ABB RAPID module: TurnProg.mod

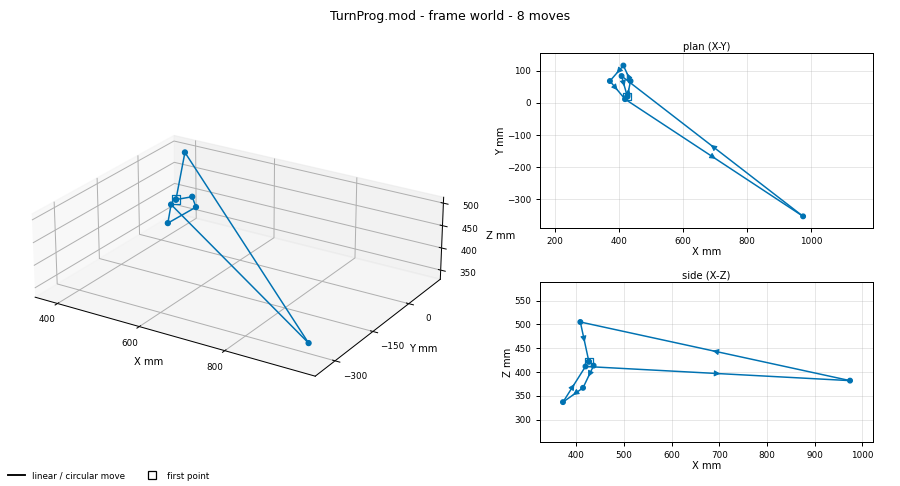
[picture p0: tool path of TurnProg.mod in frame world, 8 of 9 moves have a stored position in this frame; points joined in program order, loops and branches not executed]
%%%
  VERSION:1
  LANGUAGE:ENGLISH
%%%
MODULE MOD_TurnProg

    ! -------------------------------
    ! Define customized variables here
    ! ...

	! Tool variables:
	PERS tooldata ToolS := [TRUE,[[10.000,20.000,150.000],[1.00000000,0.00000000,0.00000000,0.00000000]],[1,[0,0,20],[1,0,0,0],0,0,0.005]];

	! Reference variables:
	PERS wobjdata FrameS := [FALSE, TRUE, "", [[0,0,0],[1,0,0,0]],[[1234.570,-98.765,50.500],[0.96592583,0.00000000,0.00000000,0.25881905]]];

	PROC Main()
		ConfJ \On;
		ConfL \Off;
		! Program generated by RoboDK v6.0.7 for ABB IRB 260 on XX/XX/XXXX 18:00:00
		! Using nominal kinematics.
		MoveL [[-640.584,506.980,371.534],[0.37410804,0.28584607,0.85365954,-0.22271191],[0,0,0,0],[9E+09,9E+09,9E+09,9E+09,9E+09,9E+09]],v500,z1,ToolS \WObj:=FrameS;
		MoveL [[-607.850,543.849,363.215],[0.37410804,0.28584607,0.85365954,-0.22271191],[0,0,0,0],[9E+09,9E+09,9E+09,9E+09,9E+09,9E+09]],v500,z1,ToolS \WObj:=FrameS;
		MoveL [[-602.951,596.788,316.595],[0.37410804,0.28584607,0.85365954,-0.22271191],[0,0,0,1],[9E+09,9E+09,9E+09,9E+09,9E+09,9E+09]],v500,z1,ToolS \WObj:=FrameS;
		MoveL [[-663.517,575.988,286.611],[0.37410804,0.28584607,0.85365954,-0.22271191],[0,0,0,4],[9E+09,9E+09,9E+09,9E+09,9E+09,9E+09]],v500,z1,ToolS \WObj:=FrameS;
		MoveL [[-650.861,503.437,361.399],[0.37410804,0.28584607,0.85365954,-0.22271191],[0,0,0,2],[9E+09,9E+09,9E+09,9E+09,9E+09,9E+09]],v500,z1,ToolS \WObj:=FrameS;
		MoveL [[-353.026,-90.135,331.702],[0.34432926,0.04805561,0.93307257,-0.09221494],[0,0,0,3],[9E+09,9E+09,9E+09,9E+09,9E+09,9E+09]],v500,z1,ToolS \WObj:=FrameS;
		MoveL [[-624.230,571.208,454.620],[0.55239178,-0.04267608,0.67304167,-0.48995609],[0,0,0,7],[9E+09,9E+09,9E+09,9E+09,9E+09,9E+09]],v500,z1,ToolS \WObj:=FrameS;
		MoveL [[-640.584,506.980,371.534],[0.37410804,0.28584607,0.85365954,-0.22271191],[0,0,0,6],[9E+09,9E+09,9E+09,9E+09,9E+09,9E+09]],v500,z1,ToolS \WObj:=FrameS;
		MoveAbsJ [[350.000000,0.000000,0.000000,-350.000000,0.000000,0.000000],[9E+09,9E+09,9E+09,9E+09,9E+09,9E+09]],v500,z1,ToolS \WObj:=FrameS;
	ENDPROC

ENDMODULE
